// TIA Portal V20 export
// export: Created 2026-10-20T12:47:02.121561Z, ExportSetting WithDefaults, DisplayName Totally Integrated Automation Portal, DisplayVersion V20 Update 6, DisplayName TIA Portal Openness, DisplayVersion V20 Update 6, DisplayName TIA Portal Version Control Interface, DisplayVersion V20 Update 6, DisplayName SINAMICS Startdrive Advanced, DisplayVersion V20 SP1, DisplayName SINAMICS Startdrive G130, G150, S120, S150, SINAMICS MV, G220, S200, S210, DisplayVersion V20 SP1, DisplayName SINAMICS Startdrive G110M, G120, G120C, G120D, G120P, G115D, DisplayVersion V20 SP1, DisplayName STEP 7 Professional, DisplayVersion V20 Update 6, DisplayName STEP 7 Safety, DisplayVersion V20 Update 2, DisplayName WinCC Basic/Comfort/Advanced, DisplayVersion V20 Update 6, DisplayName WinCC Unified, DisplayVersion V20 Update 6
FUNCTION "FindDINTFieldFragmented" : DInt   // FC20, SCL
{ S7_Optimized_Access := 'TRUE' }
VERSION : 0.1
// stored: AutoNumber true, IsIECCheckEnabled false, SetENOAutomatically false, UDAEnableTagReadback false
   VAR_INPUT
      FieldName : String;
      Str1 : String;
      Str2 : String;
   END_VAR
   VAR_TEMP
      searchStr : String;
      iStart : Int;
      iEnd : Int;
      tempVal : String;
      fieldFound : Bool;
      loopIdx : Int;
   END_VAR
BEGIN
   // Build search string
   #searchStr := CONCAT(IN1 := '"', IN2 := #FieldName);
   #searchStr := CONCAT(IN1 := #searchStr, IN2 := '" :');

   // Serach for JSON field
   #iStart := FIND(IN1 := #Str1, IN2 := #searchStr);

   IF #iStart > 0 THEN
       // Found full field in String_1
       #iEnd := FIND(IN1 := MID(IN := #Str1, P := #iStart + LEN(#searchStr), L := 20), IN2 := ',');
       IF #iEnd = 0 THEN
           #iEnd := FIND(IN1 := MID(IN := #Str1, P := #iStart + LEN(#searchStr), L := 20), IN2 := '}');
       END_IF;
       IF #iEnd > 0 THEN
           #tempVal := MID(IN := #Str1, P := #iStart + LEN(#searchStr), L := #iEnd - 1);
           #fieldFound := TRUE;
       END_IF;
   END_IF;

   // Search for full field in Str2
   IF NOT #fieldFound THEN
       #iStart := FIND(IN1 := #Str2, IN2 := #searchStr);
       IF #iStart > 0 THEN
           #iEnd := FIND(IN1 := MID(IN := #Str2, P := #iStart + LEN(#searchStr), L := 20), IN2 := ',');
           IF #iEnd = 0 THEN
               #iEnd := FIND(IN1 := MID(IN := #Str2, P := #iStart + LEN(#searchStr), L := 20), IN2 := '}');
           END_IF;
           IF #iEnd > 0 THEN
               #tempVal := MID(IN := #Str2, P := #iStart + LEN(#searchStr), L := #iEnd - 1);
               #fieldFound := TRUE;
           END_IF;
       END_IF;
   END_IF;

   // Search for fragmented field: end of name in Str1 and beginning in Str2
   IF NOT #fieldFound THEN
       // Examines last 10 characters of String_1
       FOR #loopIdx := LEN(#Str1) - 15 TO LEN(#Str1) DO
           IF MID(IN := #Str1, P := #loopIdx, L := 1) = '"' THEN
               #tempVal := MID(IN := #Str1, P := #loopIdx, L := LEN(#Str1) - #loopIdx + 1);
               #tempVal := CONCAT(IN1 := #tempVal, IN2 := #Str2); // concatenates piece from beginning of String_2
               #iStart := FIND(IN1 := #tempVal, IN2 := #searchStr);
               IF #iStart > 0 THEN
                   #iEnd := FIND(IN1 := MID(IN := #tempVal, P := #iStart + LEN(#searchStr), L := 20), IN2 := ',');
                   IF #iEnd = 0 THEN
                       #iEnd := FIND(IN1 := MID(IN := #tempVal, P := #iStart + LEN(#searchStr), L := 20), IN2 := '}');
                   END_IF;
                   IF #iEnd > 0 THEN
                       #tempVal := MID(IN := #tempVal, P := #iStart + LEN(#searchStr), L := #iEnd - 1);
                       #fieldFound := TRUE;
                   END_IF;
               END_IF;
               EXIT; // found, you can leave
           END_IF;
       END_FOR;
   END_IF;

   // Return value
   IF #fieldFound THEN
       #FindDINTFieldFragmented := STRING_TO_DINT(#tempVal);
   ELSE
       #FindDINTFieldFragmented := -9999; // default value if not found
   END_IF;
END_FUNCTION
